SUBAPPLICATION NumericValue_TO_AD2 (* VT-Eingabefeld (CInputNumber) lesen und als AD2 (bidirektional, DWORD/Bitmaske) an einen Consumer weiterreichen (z.B. AOption_AD_DEMUX_N.K). Speichert NICHT selbst - der Consumer meldet die tatsaechlich uebernommene Bitmaske ueber denselben AD2-Plug zurueck, das Echo wird auf das VT-Feld zurueckgeschrieben. *)
  (* Standard: 61499-2; Description: Copyright (c) 2026 Meisterschulen am Ostbahnhof This program and the accompanying materials are made available under the terms of the Eclipse Public License 2.0 which is available at https://www.eclipse.org/legal/epl-2.0/ SPDX-License-Identifier: EPL-2.0 *)
  (* Version 1.0, 2026-10-13, Franz Höpfinger, Meisterschulen am Ostbahnhof, DWORD/Bitmasken-Pendant zu MyLib::sys::NumericValue_TO_AUI2 - fuer AOption_AD_DEMUX_N (Multi-Select) statt AOption_AUI_DEMUX_N (Single-Select). Kein AD_TO_AUI-Zwischenschritt noetig, da AD2 bereits direkt DWORD ist. *)
  PACKAGE MyLib::sys;
  IMPORT isobus::UT::Q::const::IDs::ID_NULL;
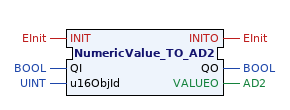
  EVENT_INPUT
    INIT : EInit; (* Initialization Request *)
  END_EVENT
  EVENT_OUTPUT
    INITO : EInit; (* Initialization Confirm *)
  END_EVENT
  VAR_INPUT
    QI : BOOL := TRUE; (* Quality Input - TRUE to enable service *)
    u16ObjId : UINT := ID_NULL; (* Object ID *)
  END_VAR
  VAR_OUTPUT
    QO : BOOL; (* Quality Output - TRUE if service executed successfully *)
  END_VAR
  PLUGS
    VALUEO : adapter::types::bidirectional::AD2;
  END_PLUGS
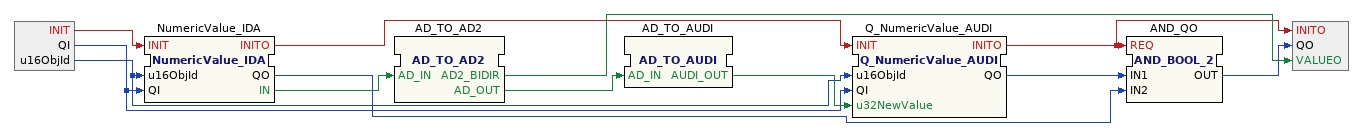
  FBS
    NumericValue_IDA : isobus::UT::io::NumericValue::NumericValue_IDA;
    AD_TO_AD2 : adapter::conversion::bidirectional::AD_TO_AD2;
    AD_TO_AUDI : adapter::conversion::unidirectional::AD_TO_AUDI;
    Q_NumericValue_AUDI : isobus::UT::Q::Q_NumericValue_AUDI;
    AND_QO : iec61131::booleanOperators::AND_BOOL_2;
  END_FBS
  EVENT_CONNECTIONS
    INIT TO NumericValue_IDA.INIT;
    NumericValue_IDA.INITO TO Q_NumericValue_AUDI.INIT;
    Q_NumericValue_AUDI.INITO TO INITO;
    Q_NumericValue_AUDI.INITO TO AND_QO.REQ;
  END_CONNECTIONS
  DATA_CONNECTIONS
    u16ObjId TO NumericValue_IDA.u16ObjId;
    u16ObjId TO Q_NumericValue_AUDI.u16ObjId;
    QI TO Q_NumericValue_AUDI.QI;
    QI TO NumericValue_IDA.QI;
    Q_NumericValue_AUDI.QO TO AND_QO.IN1;
    NumericValue_IDA.QO TO AND_QO.IN2;
    AND_QO.OUT TO QO;
  END_CONNECTIONS
  ADAPTER_CONNECTIONS
    NumericValue_IDA.IN TO AD_TO_AD2.AD_IN;
    AD_TO_AD2.AD2_BIDIR TO VALUEO;
    AD_TO_AD2.AD_OUT TO AD_TO_AUDI.AD_IN;
    AD_TO_AUDI.AUDI_OUT TO Q_NumericValue_AUDI.u32NewValue;
  END_CONNECTIONS
END_SUBAPPLICATION
